(* IEC 61131-3 sources: OpenFactory/examples/openplc, 13 files *)

(* ---- batch-mix-heat.st ---- *)
(*
  OpenFactory example PLC program: batch-mix-heat (scenes/batch-mix-heat.yaml), the batch recipe
  of PLAN 3.3: fill two ingredients to a level each, heat to a temperature, hold.
  Target: OpenPLC v3 runtime (IEC 61131-3 Structured Text), talking to the OpenFactory simulator
  as a Modbus TCP Slave Device. Setup: docs/guides/openplc-quickstart.md, then
  docs/guides/batch-mix-heat.md for this scene.

  Training and demo use only. Not a safety-rated program and not a safety-rated simulation.

  Sequence of operations (one batch, then held); BATCH_STEP holds the active step
    0.  Idle: wait 1 s after power-up for the transmitters' first readings, then start a batch
        if the mixing tank is empty (level below 0.02 m).
    10. Fill water: open XV_01 until the level reaches 0.10 m.
    20. Fill syrup: open XV_02 until the level reaches 0.16 m (the recipe: 0.06 m of syrup on
        0.10 m of water, 37.5 % syrup by volume; each valve's 1 s close adds a little).
    30. Heat: the heater runs until the temperature reaches 50 C.
    40. Hold: the batch is ready (PL_READY_DO lit); the heater keeps it at 50 C, on below
        49.5 C and off at 50 C.
    Interlocks, in every step: the high level switch (LSH) closes both inlet valves, and the
    heater runs only while the level covers it (0.10 m and above).

  I/O map: Modbus addresses come from the scene's int16_scaled lockfile
  (scenes/batch-mix-heat.int16_scaled.modbus.yaml) and the exported I/O list CSV. OpenPLC places
  a Slave Device's points from address 100 onward, so a zero-based Modbus address N maps to
  %IX100.N, %QX100.N or %IW100+N.
*)
PROGRAM batch_mix_heat
  VAR
    (* Discrete inputs from the simulator (Modbus DI:0..3) *)
    TK_01_LSH_DI AT %IX100.0 : BOOL;    (* DI:0 Batch Mixing Tank - high level switch (LSH), 0.5 m *)
    XV_01_ZSC_DI AT %IX100.1 : BOOL;    (* DI:1 Mixing Tank Water Inlet Valve - closed limit (ZSC) *)
    XV_02_ZSC_DI AT %IX100.2 : BOOL;    (* DI:2 Mixing Tank Syrup Inlet Valve - closed limit (ZSC) *)
    SIM_HEARTBEAT_DI AT %IX100.3 : BOOL; (* DI:3 OpenFactory simulator heartbeat, 1 Hz; not used here, watch it for a sim-down watchdog *)
    (* Coils to the simulator (Modbus CO:0..3) *)
    HTR_01_ON_DO AT %QX100.0 : BOOL;    (* CO:0 Batch Mixing Tank Immersion Heater - on command *)
    PL_READY_DO AT %QX100.1 : BOOL;     (* CO:1 Batch Ready Pilot Light *)
    XV_01_OPEN_DO AT %QX100.2 : BOOL;   (* CO:2 Mixing Tank Water Inlet Valve - open command *)
    XV_02_OPEN_DO AT %QX100.3 : BOOL;   (* CO:3 Mixing Tank Syrup Inlet Valve - open command *)
    (* Input registers (Modbus IR:0..1) *)
    TK_01_LT_AI AT %IW100 : INT;        (* IR:0 Batch Mixing Tank Level Transmitter, 0 to 32767 = 0 to 0.6 m *)
    TK_01_TT_AI AT %IW101 : INT;        (* IR:1 Batch Mixing Tank Temperature Transmitter, 0 to 32767 = 0 to 100 C *)
  END_VAR
  VAR
    WATER_SP : REAL := 0.10;            (* level at which the water fill ends, m *)
    BATCH_SP : REAL := 0.16;            (* level at which the syrup fill ends, m *)
    EMPTY_LVL : REAL := 0.02;           (* below this the tank is empty and can start a batch, m *)
    TEMP_SP : REAL := 50.0;             (* batch temperature, C *)
    HOLD_DB : REAL := 0.5;              (* the heater restarts this far below TEMP_SP in the hold, C *)
    COVER_LVL : REAL := 0.10;           (* heater low-level permissive, m *)
    STARTUP_DELAY : TIME := T#1s;       (* until the transmitters' first readings *)
    STARTUP_TMR : TON;
    BATCH_STEP : INT := 0;              (* the active step: 0, 10, 20, 30, 40; not STEP, an IEC 61131-3 keyword *)
    HEAT : BOOL := FALSE;               (* heater demand before the permissive *)
    LEVEL_M : REAL;
    TEMP_C : REAL;
  END_VAR

  LEVEL_M := INT_TO_REAL(TK_01_LT_AI) * 0.6 / 32767.0;
  TEMP_C := INT_TO_REAL(TK_01_TT_AI) * 100.0 / 32767.0;
  STARTUP_TMR(IN := TRUE, PT := STARTUP_DELAY);

  (* Transitions, one per scan *)
  CASE BATCH_STEP OF
    0:  IF STARTUP_TMR.Q AND LEVEL_M < EMPTY_LVL THEN BATCH_STEP := 10; END_IF;
    10: IF LEVEL_M >= WATER_SP THEN BATCH_STEP := 20; END_IF;
    20: IF LEVEL_M >= BATCH_SP THEN BATCH_STEP := 30; END_IF;
    30: IF TEMP_C >= TEMP_SP THEN BATCH_STEP := 40; END_IF;
  END_CASE;

  (* Actions; the hold is a thermostat with a deadband *)
  IF BATCH_STEP = 30 THEN
    HEAT := TRUE;
  ELSIF BATCH_STEP = 40 THEN
    IF TEMP_C >= TEMP_SP THEN
      HEAT := FALSE;
    ELSIF TEMP_C < TEMP_SP - HOLD_DB THEN
      HEAT := TRUE;
    END_IF;
  ELSE
    HEAT := FALSE;
  END_IF;
  XV_01_OPEN_DO := (BATCH_STEP = 10) AND NOT TK_01_LSH_DI;
  XV_02_OPEN_DO := (BATCH_STEP = 20) AND NOT TK_01_LSH_DI;
  HTR_01_ON_DO := HEAT AND LEVEL_M >= COVER_LVL;
  PL_READY_DO := (BATCH_STEP = 40);
END_PROGRAM

CONFIGURATION Config0
  RESOURCE Res0 ON PLC
    TASK task0(INTERVAL := T#20ms, PRIORITY := 0);
    PROGRAM instance0 WITH task0 : batch_mix_heat;
  END_RESOURCE
END_CONFIGURATION

(* ---- buffer-and-release.st ---- *)
(*
  OpenFactory example PLC program: buffer-and-release (scenes/buffer-and-release.yaml), PLAN 2.7.
  Target: OpenPLC v3 runtime (IEC 61131-3 Structured Text), talking to the OpenFactory simulator
  as a Modbus TCP Slave Device. Setup: docs/guides/openplc-quickstart.md, then
  docs/guides/buffer-and-release.md for this scene.

  Training and demo use only. Not a safety-rated program and not a safety-rated simulation.

  Sequence of operations
    1. Run both belts. Hold STP_01 raised, so boxes queue nose to tail on the buffer belt.
    2. Enable the box emitter once both belts have reported running for 1 s.
    3. A batch is ready when PE_FULL (under the third queued box) has been blocked for 1.5 s, which
       a moving box (1 s in the beam at 0.3 m/s) cannot do, and the blade has been back up for at
       least 2 s since the last batch.
    4. Release: lower STP_01 and count PE_REL rising edges on the outfeed belt. The outfeed runs
       three times faster than the buffer, so each released box pulls a gap and the eye clears
       between boxes. At the third, raise the blade: the fourth box is still behind the blade line.

  Timing margin: when the third box of a batch reaches PE_REL, the fourth box's front is about
  0.10 m behind the blade line, 0.33 s at 0.3 m/s. OpenPLC sees the eye up to 100 ms late and
  writes the raise up to 100 ms later, which that margin covers. The blade holds parts from the
  moment it starts rising; a box already over the blade line passes.

  I/O map: Modbus addresses come from the scene's int16_scaled lockfile
  (scenes/buffer-and-release.int16_scaled.modbus.yaml) and the exported I/O list CSV. OpenPLC
  places a Slave Device's points from address 100 onward, so a zero-based Modbus address N maps
  to %IX100.N or %QX100.N. The scene has no analog tags, so both lockfiles give the same addresses.
*)
PROGRAM buffer_release
  VAR
    (* Discrete inputs from the simulator (Modbus DI:0..6) *)
    CONV_BUF_RUN_DI AT %IX100.0 : BOOL; (* DI:0 Buffer Belt Conveyor - running feedback *)
    CONV_OUT_RUN_DI AT %IX100.1 : BOOL; (* DI:1 Outfeed Belt Conveyor - running feedback *)
    PE_FULL_DI AT %IX100.2 : BOOL;      (* DI:2 Buffer Batch Ready Photo Eye - beam blocked *)
    PE_REL_DI AT %IX100.3 : BOOL;       (* DI:3 Outfeed Release Count Photo Eye - beam blocked *)
    STP_01_DN_DI AT %IX100.4 : BOOL;    (* DI:4 Buffer Release Stopper - lowered limit *)
    STP_01_UP_DI AT %IX100.5 : BOOL;    (* DI:5 Buffer Release Stopper - raised limit *)
    SIM_HEARTBEAT_DI AT %IX100.6 : BOOL; (* DI:6 OpenFactory simulator heartbeat, 1 Hz; not used here, watch it for a sim-down watchdog *)
    (* Coils to the simulator (Modbus CO:0..3) *)
    CONV_BUF_RUN_DO AT %QX100.0 : BOOL; (* CO:0 Buffer Belt Conveyor - run command *)
    CONV_OUT_RUN_DO AT %QX100.1 : BOOL; (* CO:1 Outfeed Belt Conveyor - run command *)
    EMT_01_EN_DO AT %QX100.2 : BOOL;    (* CO:2 Buffer Belt Box Source - enable *)
    STP_01_RAISE_DO AT %QX100.3 : BOOL; (* CO:3 Buffer Release Stopper - raise solenoid *)
  END_VAR
  VAR
    BATCH : INT := 3;                   (* boxes per release *)
    BELTS_OK_DELAY : TIME := T#1s;      (* run feedback must hold this long to feed boxes *)
    FULL_DELAY : TIME := T#1500ms;      (* a standing box, not a passing one, at PE_FULL *)
    PAUSE : TIME := T#2s;               (* blade up at least this long between batches *)
    BELTS_OK_TMR : TON;                 (* both belts running, debounced *)
    FULL_TMR : TON;                     (* a box stands under PE_FULL: three are queued *)
    PAUSE_TMR : TON;                    (* the blade has been back up PAUSE since the last batch *)
    PE_REL_RISE : R_TRIG;               (* a released box reaches PE_REL *)
    RELEASING : BOOL;                   (* a batch is on its way out *)
    RELEASED : INT;                     (* boxes counted out in this batch *)
  END_VAR

  (* 1. Belts run *)
  CONV_BUF_RUN_DO := TRUE;
  CONV_OUT_RUN_DO := TRUE;

  (* 2. Feed boxes only after both belts have reported running for BELTS_OK_DELAY *)
  BELTS_OK_TMR(IN := CONV_BUF_RUN_DI AND CONV_OUT_RUN_DI, PT := BELTS_OK_DELAY);
  EMT_01_EN_DO := BELTS_OK_TMR.Q;

  (* 3. A batch is ready: three queued, and the blade up long enough since the last batch *)
  FULL_TMR(IN := PE_FULL_DI, PT := FULL_DELAY);
  PAUSE_TMR(IN := STP_01_UP_DI AND NOT RELEASING, PT := PAUSE);
  IF FULL_TMR.Q AND PAUSE_TMR.Q AND NOT RELEASING THEN
    RELEASING := TRUE;
    RELEASED := 0;
  END_IF;

  (* 4. Count the batch out on the outfeed; raise the blade at the last one *)
  PE_REL_RISE(CLK := PE_REL_DI);
  IF PE_REL_RISE.Q AND RELEASING THEN
    RELEASED := RELEASED + 1;
    IF RELEASED >= BATCH THEN
      RELEASING := FALSE;
    END_IF;
  END_IF;
  STP_01_RAISE_DO := NOT RELEASING;
END_PROGRAM

CONFIGURATION Config0
  RESOURCE Res0 ON PLC
    TASK task0(INTERVAL := T#20ms, PRIORITY := 0);
    PROGRAM instance0 WITH task0 : buffer_release;
  END_RESOURCE
END_CONFIGURATION

(* ---- conveyor-start-stop.st ---- *)
(*
  OpenFactory example PLC program: conveyor-start-stop (scenes/conveyor-start-stop.yaml), the
  hello-world scene of PLAN 2.7.
  Target: OpenPLC v3 runtime (IEC 61131-3 Structured Text), talking to the OpenFactory simulator
  as a Modbus TCP Slave Device. Setup: docs/guides/openplc-quickstart.md, then
  docs/guides/conveyor-start-stop.md for this scene.

  Training and demo use only. Not a safety-rated program and not a safety-rated simulation.
  A real stop circuit is hard-wired; a PLC stop input like this one is an operator convenience.

  Sequence of operations
    1. Turning SS_01 to RUN starts the line: CONV_01 runs and stays running (seal-in) while SS_01
       stays in RUN and PB_STOP is not pressed. The scene starts with SS_01 in RUN, so the line
       starts on the first scan that sees it there.
    2. PB_STOP is wired normally closed (the scene binds it with invert: true): PB_STOP_DI is TRUE
       while the button is released, and a broken wire reads as a press, so it fails safe.
       Pressing it drops the seal-in. To restart, turn SS_01 to OFF and back to RUN.
    3. A selector reading OFF and RUN at once (a wiring fault) stops the line too.
    4. Once CONV_01 has reported running for 1 s, enable the box emitter EMT_01.
    5. PL_RUN shows the running feedback, not the command.
    Boxes ride the belt end to end and reach REM_01.

  I/O map: Modbus addresses come from the scene's int16_scaled lockfile
  (scenes/conveyor-start-stop.int16_scaled.modbus.yaml) and the exported I/O list CSV. OpenPLC
  places a Slave Device's points from address 100 onward, so a zero-based Modbus address N maps to
  %IX100.N or %QX100.N. This scene has no analog tags, so the float32 and int16_scaled lockfiles
  give the same addresses (ADR-0004 decision 8).

  Why the emitter waits 1 s: see examples/openplc/sorting-by-height.st. When OpenPLC (re)connects,
  its input image can hold old feedback for one poll, and an enable written straight from it can
  chatter and drop two boxes on top of each other.
*)
PROGRAM start_stop
  VAR
    (* Discrete inputs from the simulator (Modbus DI:0..4) *)
    CONV_01_RUN_DI AT %IX100.0 : BOOL;  (* DI:0 Transfer Belt Conveyor - running feedback *)
    PB_STOP_DI AT %IX100.1 : BOOL;      (* DI:1 Transfer Conveyor Stop Pushbutton - NC, TRUE = released *)
    SS_01_OFF_DI AT %IX100.2 : BOOL;    (* DI:2 Off/Run Selector Switch - in OFF *)
    SS_01_RUN_DI AT %IX100.3 : BOOL;    (* DI:3 Off/Run Selector Switch - in RUN *)
    SIM_HEARTBEAT_DI AT %IX100.4 : BOOL; (* DI:4 OpenFactory simulator heartbeat, 1 Hz; not used here, watch it for a sim-down watchdog *)
    (* Coils to the simulator (Modbus CO:0..2) *)
    CONV_01_RUN_DO AT %QX100.0 : BOOL;  (* CO:0 Transfer Belt Conveyor - run command *)
    EMT_01_EN_DO AT %QX100.1 : BOOL;    (* CO:1 Transfer Belt Box Source - enable *)
    PL_RUN_DO AT %QX100.2 : BOOL;       (* CO:2 Transfer Conveyor Running Pilot Light *)
  END_VAR
  VAR
    BELT_OK_DELAY : TIME := T#1s;       (* running feedback must hold this long to feed boxes *)
    BELT_OK_TMR : TON;                  (* belt running, debounced *)
    SS_RUN_RISE : R_TRIG;               (* selector turned to RUN (also the first scan in RUN) *)
    RUN_OK : BOOL;                      (* selector in RUN only, stop button released *)
    RUN_LATCH : BOOL;                   (* the line is started (seal-in) *)
  END_VAR

  (* 1-3. Start on a turn to RUN, seal in, drop on stop, OFF, or a selector wiring fault *)
  RUN_OK := SS_01_RUN_DI AND NOT SS_01_OFF_DI AND PB_STOP_DI;
  SS_RUN_RISE(CLK := SS_01_RUN_DI);
  RUN_LATCH := (SS_RUN_RISE.Q OR RUN_LATCH) AND RUN_OK;
  CONV_01_RUN_DO := RUN_LATCH;

  (* 4. Feed boxes only after the belt has reported running for BELT_OK_DELAY *)
  BELT_OK_TMR(IN := RUN_LATCH AND CONV_01_RUN_DI, PT := BELT_OK_DELAY);
  EMT_01_EN_DO := BELT_OK_TMR.Q;

  (* 5. Running light from feedback *)
  PL_RUN_DO := CONV_01_RUN_DI;
END_PROGRAM

CONFIGURATION Config0
  RESOURCE Res0 ON PLC
    TASK task0(INTERVAL := T#20ms, PRIORITY := 0);
    PROGRAM instance0 WITH task0 : start_stop;
  END_RESOURCE
END_CONFIGURATION

(* ---- inline-reject.st ---- *)
(*
  OpenFactory example PLC program: inline-reject (scenes/inline-reject.yaml).
  Target: OpenPLC v3 runtime (IEC 61131-3 Structured Text), talking to the OpenFactory simulator
  as a Modbus TCP Slave Device. Setup: docs/guides/openplc-quickstart.md.

  Training and demo use only. Not a safety-rated program and not a safety-rated simulation.

  The scene was built in the scene editor from `openfactory new`, without the file being opened
  (docs/guides/inline-reject.md). This program is a line-for-line port of the stand-in script,
  examples/pyplc/inline-reject.py.

  Sequence of operations
    1. Run both belt conveyors (CONV_01 feeds CONV_02 end to end).
    2. Enable the box emitter once both belts have reported running for 1 s without a break.
    3. PE_01 sits 0.3 m above CONV_02: oversize boxes (0.4 m) break the beam, good ones (0.2 m)
       pass under it. On each PE_01 rising edge, start that box's own REJECT_DELAY timer for its
       travel from the eye to the pusher plate, then extend CYL_01 when it expires; the plate
       pushes the box off the side of CONV_02 into the reject bin, REM_01. Each oversize box
       takes the next of four slots (a ring: REJECT_PEND_n and REJECT_TMR_n).
    4. Retract CYL_01 as soon as its extended limit (CYL_01_EXTENDED_DI) is made.
    Good boxes ride on to the end of CONV_02 and reach REM_02.

  I/O map: Modbus addresses come from the scene's lockfiles (scenes/inline-reject.*.modbus.yaml;
  this scene has no analog tags, so both give the same addresses). OpenPLC places a Slave
  Device's points from address 100 onward, so a zero-based Modbus address N maps to %IX100.N or
  %QX100.N.

  Timing: the eye and the plate are 1.0 m apart along CONV_02, as on sorting-by-height, so the
  box is due at the plate 2.08 s after it trips the eye at 0.5 m/s; REJECT_DELAY is 2.08 s minus
  OpenPLC's average 0.10 s polling latency, as the sorter's DIVERT_DELAY is.
*)
PROGRAM inline_reject
  VAR
    (* Discrete inputs from the simulator (Modbus DI:0..4) *)
    CONV_01_RUNNING_DI AT %IX100.0 : BOOL;  (* DI:0 Infeed Belt Conveyor - running feedback *)
    CONV_02_RUNNING_DI AT %IX100.1 : BOOL;  (* DI:1 Outfeed Belt Conveyor - running feedback *)
    CYL_01_EXTENDED_DI AT %IX100.2 : BOOL;  (* DI:2 Oversize Box Reject Pusher - extended limit *)
    PE_01_DI AT %IX100.3 : BOOL;            (* DI:3 Oversize Box Photo Eye - beam blocked *)
    SIM_HEARTBEAT_DI AT %IX100.4 : BOOL;    (* DI:4 OpenFactory simulator heartbeat, 1 Hz; not used here *)
    (* Coils to the simulator (Modbus CO:0..3) *)
    CONV_01_RUN_DO AT %QX100.0 : BOOL;      (* CO:0 Infeed Belt Conveyor - run command *)
    CONV_02_RUN_DO AT %QX100.1 : BOOL;      (* CO:1 Outfeed Belt Conveyor - run command *)
    CYL_01_EXTEND_DO AT %QX100.2 : BOOL;    (* CO:2 Oversize Box Reject Pusher - extend solenoid *)
    EMT_01_DO AT %QX100.3 : BOOL;           (* CO:3 Infeed Box Source - enable *)
  END_VAR
  VAR
    REJECT_DELAY : TIME := T#1980ms;    (* eye-to-plate travel, less average polling latency *)
    BELTS_OK_DELAY : TIME := T#1s;      (* run feedback must hold this long to feed boxes *)
    BELTS_OK_TMR : TON;                 (* both belts running, debounced *)
    PE_01_RISE : R_TRIG;                (* an oversize box arrives at PE_01 *)
    REJECT_TMR_0 : TON;                 (* eye-to-plate travel timer, slot 0 *)
    REJECT_TMR_1 : TON;                 (* eye-to-plate travel timer, slot 1 *)
    REJECT_TMR_2 : TON;                 (* eye-to-plate travel timer, slot 2 *)
    REJECT_TMR_3 : TON;                 (* eye-to-plate travel timer, slot 3 *)
    REJECT_PEND_0 : BOOL;               (* slot 0 holds an oversize box on its way to the pusher *)
    REJECT_PEND_1 : BOOL;               (* slot 1 holds an oversize box on its way to the pusher *)
    REJECT_PEND_2 : BOOL;               (* slot 2 holds an oversize box on its way to the pusher *)
    REJECT_PEND_3 : BOOL;               (* slot 3 holds an oversize box on its way to the pusher *)
    NEXT_SLOT : INT := 0;               (* ring index: the slot the next oversize box takes, 0..3 *)
    PUSH_CMD : BOOL;                    (* pusher extend request, held until the extended limit *)
  END_VAR

  (* 1. Belts run *)
  CONV_01_RUN_DO := TRUE;
  CONV_02_RUN_DO := TRUE;

  (* 2. Feed boxes only after both belts have reported running for BELTS_OK_DELAY *)
  BELTS_OK_TMR(IN := CONV_01_RUNNING_DI AND CONV_02_RUNNING_DI, PT := BELTS_OK_DELAY);
  EMT_01_DO := BELTS_OK_TMR.Q;

  (* 3. Oversize box at the eye: give it the next slot and its own travel timer *)
  PE_01_RISE(CLK := PE_01_DI);
  IF PE_01_RISE.Q THEN
    CASE NEXT_SLOT OF
      0: REJECT_PEND_0 := TRUE;
      1: REJECT_PEND_1 := TRUE;
      2: REJECT_PEND_2 := TRUE;
      3: REJECT_PEND_3 := TRUE;
    END_CASE;
    NEXT_SLOT := (NEXT_SLOT + 1) MOD 4;
  END_IF;

  (* 3a. Each slot's box is due at the plate: extend *)
  REJECT_TMR_0(IN := REJECT_PEND_0, PT := REJECT_DELAY);
  IF REJECT_TMR_0.Q THEN
    REJECT_PEND_0 := FALSE;
    PUSH_CMD := TRUE;
  END_IF;
  REJECT_TMR_1(IN := REJECT_PEND_1, PT := REJECT_DELAY);
  IF REJECT_TMR_1.Q THEN
    REJECT_PEND_1 := FALSE;
    PUSH_CMD := TRUE;
  END_IF;
  REJECT_TMR_2(IN := REJECT_PEND_2, PT := REJECT_DELAY);
  IF REJECT_TMR_2.Q THEN
    REJECT_PEND_2 := FALSE;
    PUSH_CMD := TRUE;
  END_IF;
  REJECT_TMR_3(IN := REJECT_PEND_3, PT := REJECT_DELAY);
  IF REJECT_TMR_3.Q THEN
    REJECT_PEND_3 := FALSE;
    PUSH_CMD := TRUE;
  END_IF;

  (* 4. Retract on the extended limit *)
  IF CYL_01_EXTENDED_DI THEN
    PUSH_CMD := FALSE;
  END_IF;
  CYL_01_EXTEND_DO := PUSH_CMD;
END_PROGRAM

CONFIGURATION Config0
  RESOURCE Res0 ON PLC
    TASK task0(INTERVAL := T#20ms, PRIORITY := 0);
    PROGRAM instance0 WITH task0 : inline_reject;
  END_RESOURCE
END_CONFIGURATION

(* ---- palletizer-lite.st ---- *)
(*
  OpenFactory example PLC program: palletizer-lite (scenes/palletizer-lite.yaml), PLAN 2.7.
  Target: OpenPLC v3 runtime (IEC 61131-3 Structured Text), talking to the OpenFactory simulator
  as a Modbus TCP Slave Device. Setup: docs/guides/openplc-quickstart.md, then
  docs/guides/palletizer-lite.md for this scene.

  Training and demo use only. Not a safety-rated program and not a safety-rated simulation.

  Sequence of operations
    1. Run both belts and hold both stoppers raised; enable the box source once both belts have
       reported running for 1 s. Boxes queue at STP_IN, the first one under the gantry.
    2. Pick and place, one box per cycle (the gantry has no raised switch, so each rise is timed):
       with a box at PE_PICK, the gantry at the pick side, fewer than LAYER_BOXES placed in this
       layer, and no layer leaving: PICK_STEP 1 lower, 2 grip, 3 rise, 4 traverse, 5 lower,
       6 release, 7 rise, 8 return, back to 0. (STEP is a reserved word in IEC 61131-3.) Count each box placed. The layer-forming belt carries it to
       the row queueing at STP_LYR.
    3. A layer is complete when LAYER_BOXES have been placed and PE_ROW (under the fourth queued
       box) has been blocked for 1 s, which a passing box (0.6 s in the beam) cannot do. Lower
       STP_LYR for LAYER_OUT to send the layer to the discharge, raise it, and start the count
       again. Counting placements, not just watching PE_ROW, keeps a fifth box from being set
       down while the row completes and riding out with the layer.

  I/O map: Modbus addresses come from the scene's int16_scaled lockfile
  (scenes/palletizer-lite.int16_scaled.modbus.yaml) and the exported I/O list CSV. OpenPLC places
  a Slave Device's points from address 100 onward, eight bits to a byte: zero-based Modbus address
  N maps to %IX(100 + N / 8).(N MOD 8), and likewise for %QX. The scene has no analog tags, so
  both lockfiles give the same addresses.
*)
PROGRAM palletizer
  VAR
    (* Discrete inputs from the simulator (Modbus DI:0..8) *)
    CONV_IN_RUN_DI AT %IX100.0 : BOOL;  (* DI:0 Palletizer Infeed Belt Conveyor - running *)
    CONV_LYR_RUN_DI AT %IX100.1 : BOOL; (* DI:1 Layer Forming Belt Conveyor - running *)
    PE_PICK_DI AT %IX100.2 : BOOL;      (* DI:2 Infeed Box At Pick Position Photo Eye *)
    PE_ROW_DI AT %IX100.3 : BOOL;       (* DI:3 Layer Row Complete Photo Eye *)
    PP_01_AT_PICK_DI AT %IX100.4 : BOOL;  (* DI:4 Transfer Gantry - at pick side *)
    PP_01_AT_PLACE_DI AT %IX100.5 : BOOL; (* DI:5 Transfer Gantry - at place side *)
    PP_01_DOWN_DI AT %IX100.6 : BOOL;   (* DI:6 Transfer Gantry - pad lowered *)
    PP_01_HOLD_DI AT %IX100.7 : BOOL;   (* DI:7 Transfer Gantry - holding a part *)
    SIM_HEARTBEAT_DI AT %IX100.8 : BOOL; (* DI:8 OpenFactory simulator heartbeat, 1 Hz; not used here, watch it for a sim-down watchdog *)
    (* Coils to the simulator (Modbus CO:0..7) *)
    CONV_IN_RUN_DO AT %QX100.0 : BOOL;  (* CO:0 Palletizer Infeed Belt Conveyor - run *)
    CONV_LYR_RUN_DO AT %QX100.1 : BOOL; (* CO:1 Layer Forming Belt Conveyor - run *)
    EMT_01_EN_DO AT %QX100.2 : BOOL;    (* CO:2 Palletizer Infeed Box Source - enable *)
    PP_01_GRIP_DO AT %QX100.3 : BOOL;   (* CO:3 Transfer Gantry - grip *)
    PP_01_LOWER_DO AT %QX100.4 : BOOL;  (* CO:4 Transfer Gantry - lower pad *)
    PP_01_TRAV_DO AT %QX100.5 : BOOL;   (* CO:5 Transfer Gantry - traverse to place side *)
    STP_IN_RAISE_DO AT %QX100.6 : BOOL; (* CO:6 Infeed Pick Position Stopper - raise *)
    STP_LYR_RAISE_DO AT %QX100.7 : BOOL; (* CO:7 Layer Forming Stopper - raise *)
  END_VAR
  VAR
    LAYER_BOXES : INT := 4;             (* boxes per layer *)
    BELTS_OK_DELAY : TIME := T#1s;      (* run feedback must hold this long to feed boxes *)
    RISE : TIME := T#400ms;             (* pad rise, lower_time_s 0.3 plus margin *)
    SETTLE : TIME := T#200ms;           (* the released box drops onto the belt *)
    ROW_DELAY : TIME := T#1s;           (* a standing box, not a passing one, at PE_ROW *)
    LAYER_OUT : TIME := T#3s;           (* four boxes (1.2 m) clear the blade at 0.5 m/s *)
    BELTS_OK_TMR : TON;                 (* both belts running, debounced *)
    RISE_TMR : TON;                     (* the pad has had time to rise *)
    SETTLE_TMR : TON;                   (* the released box has settled on the belt *)
    ROW_TMR : TON;                      (* a box stands under PE_ROW *)
    LAYER_TMR : TON;                    (* the layer has had time to leave *)
    PICK_STEP : INT := 0;               (* pick-and-place step, 0 = waiting at the pick side *)
    LAYER_OUT_ON : BOOL;                (* a layer is leaving *)
    PLACED : INT := 0;                  (* boxes placed in the layer being formed *)
  END_VAR

  (* 1. Belts run; stoppers hold; feed boxes once both belts report running for 1 s *)
  CONV_IN_RUN_DO := TRUE;
  CONV_LYR_RUN_DO := TRUE;
  STP_IN_RAISE_DO := TRUE;
  BELTS_OK_TMR(IN := CONV_IN_RUN_DI AND CONV_LYR_RUN_DI, PT := BELTS_OK_DELAY);
  EMT_01_EN_DO := BELTS_OK_TMR.Q;

  (* 2. Pick and place, one box per cycle; the timers run only in the steps that use them *)
  RISE_TMR(IN := PICK_STEP = 3 OR PICK_STEP = 7, PT := RISE);
  SETTLE_TMR(IN := PICK_STEP = 6 AND NOT PP_01_HOLD_DI, PT := SETTLE);
  CASE PICK_STEP OF
    0: IF PE_PICK_DI AND PP_01_AT_PICK_DI AND PLACED < LAYER_BOXES AND NOT LAYER_OUT_ON THEN
         PICK_STEP := 1;
       END_IF;
    1: IF PP_01_DOWN_DI THEN PICK_STEP := 2; END_IF;
    2: IF PP_01_HOLD_DI THEN PICK_STEP := 3; END_IF;
    3: IF RISE_TMR.Q THEN PICK_STEP := 4; END_IF;
    4: IF PP_01_AT_PLACE_DI THEN PICK_STEP := 5; END_IF;
    5: IF PP_01_DOWN_DI THEN PICK_STEP := 6; END_IF;
    6: IF SETTLE_TMR.Q THEN
         PICK_STEP := 7;
         PLACED := PLACED + 1;
       END_IF;
    7: IF RISE_TMR.Q THEN PICK_STEP := 8; END_IF;
    8: IF PP_01_AT_PICK_DI THEN PICK_STEP := 0; END_IF;
  END_CASE;
  PP_01_LOWER_DO := PICK_STEP = 1 OR PICK_STEP = 2 OR PICK_STEP = 5 OR PICK_STEP = 6;
  PP_01_GRIP_DO := PICK_STEP = 2 OR PICK_STEP = 3 OR PICK_STEP = 4 OR PICK_STEP = 5;
  PP_01_TRAV_DO := PICK_STEP = 4 OR PICK_STEP = 5 OR PICK_STEP = 6 OR PICK_STEP = 7;

  (* 3. A complete row leaves as one layer *)
  ROW_TMR(IN := PE_ROW_DI, PT := ROW_DELAY);
  IF ROW_TMR.Q AND PLACED >= LAYER_BOXES AND NOT LAYER_OUT_ON THEN
    LAYER_OUT_ON := TRUE;
  END_IF;
  LAYER_TMR(IN := LAYER_OUT_ON, PT := LAYER_OUT);
  IF LAYER_TMR.Q THEN
    LAYER_OUT_ON := FALSE;
    PLACED := 0;
  END_IF;
  STP_LYR_RAISE_DO := NOT LAYER_OUT_ON;
END_PROGRAM

CONFIGURATION Config0
  RESOURCE Res0 ON PLC
    TASK task0(INTERVAL := T#20ms, PRIORITY := 0);
    PROGRAM instance0 WITH task0 : palletizer;
  END_RESOURCE
END_CONFIGURATION

(* ---- plantpax-tank-level.st ---- *)
(*
  OpenFactory example PLC program: plantpax-tank-level (scenes/plantpax-tank-level.yaml), the
  PlantPAx demo plant of PLAN 3.4 controlled without PlantPAx: tank-level-pid's level loop closed
  with OpenPLC's PID function block, plus the transfer pump. The PlantPAx version of the same
  control is the L5X from `openfactory export ... --format plantpax` (docs/plantpax.md).
  Target: OpenPLC v3 runtime (IEC 61131-3 Structured Text), talking to the OpenFactory simulator
  as a Modbus TCP Slave Device. Setup: docs/guides/openplc-quickstart.md, then
  docs/guides/plantpax-tank-level.md for this scene.

  Training and demo use only. Not a safety-rated program and not a safety-rated simulation.

  The PID block is the one in OpenPLC's compiler library (matiec lib/pid_st.txt, from the IEC
  61131-3 2nd edition draft): XOUT := KP * (ERROR + ITERM.XOUT / TR + DTERM.XOUT * TD) with
  ERROR := PV - SP. The error is PV minus SP, so a loop that opens the inlet valve on a low level
  needs a negative KP. Its integral (lib/integral_st.txt) is a rectangular sum of ERROR times
  TIME_TO_REAL(CYCLE). It has no output limit and no anti-windup: LIMIT clamps the output here,
  and the interlock holds the block in manual so it cannot wind up while overridden.
  [TBD: verify on the first OpenPLC run] that TIME_TO_REAL(T#20ms) is 0.02 (seconds) in the
  runtime; the gains below assume seconds, as the stand-in script does.

  Sequence of operations
    1. Read the level from the transmitter, raw 0 to 32767 for 0 to 2 m.
    2. PI control: the valve position is KP * (e + sum(e * 0.02 s) / TR) with e = level - 1.0 m.
    3. The output is limited to 0 to 100 % and written to the valve, raw 0 to 32767.
    4. Interlock: while the high level switch (LSH) is on, the valve is closed and the PID is
       held in manual at 0 % (no windup while it is overridden).
    5. For the first second the PID runs in manual at the valve's starting position (66 %),
       tracking the level, then switches to automatic bumplessly: the level input reads 0 until
       its first poll, and starting in automatic on that would slam the valve shut.
    6. The transfer pump P_01 starts 20 s after power-up (the demo's load step) and runs while
       the low level switch (LSL) is off: LSL is its interlock against running the tank dry.

  I/O map: Modbus addresses come from the scene's int16_scaled lockfile
  (scenes/plantpax-tank-level.int16_scaled.modbus.yaml) and the exported I/O list CSV. OpenPLC places
  a Slave Device's points from address 100 onward, so a zero-based Modbus address N maps to
  %IX100.N, %IW100+N, or %QW100+N.
*)
PROGRAM plantpax_tank
  VAR
    (* Discrete inputs from the simulator (Modbus DI:0..3) *)
    P_01_RUN_DI AT %IX100.0 : BOOL;     (* DI:0 Level Control Tank Transfer Pump - running feedback *)
    TK_01_LSH_DI AT %IX100.1 : BOOL;    (* DI:1 Level Control Tank - high level switch (LSH), 1.8 m *)
    TK_01_LSL_DI AT %IX100.2 : BOOL;    (* DI:2 Level Control Tank - low level switch (LSL), 0.3 m *)
    SIM_HEARTBEAT_DI AT %IX100.3 : BOOL; (* DI:3 OpenFactory simulator heartbeat, 1 Hz; not used here, watch it for a sim-down watchdog *)
    (* Coils to the simulator (Modbus CO:0) *)
    P_01_RUN_DO AT %QX100.0 : BOOL;     (* CO:0 Level Control Tank Transfer Pump - run command *)
    (* Input registers (Modbus IR:0..1) *)
    FV_01_ZT_AI AT %IW100 : INT;        (* IR:0 Tank Inlet Level Control Valve - position feedback, 0 to 32767 = 0 to 100 % *)
    TK_01_LT_AI AT %IW101 : INT;        (* IR:1 Level Control Tank Level Transmitter, 0 to 32767 = 0 to 2 m *)
    (* Holding registers to the simulator (Modbus HR:0) *)
    FV_01_POS_AO AT %QW100 : INT;       (* HR:0 Tank Inlet Level Control Valve - position command, 0 to 32767 = 0 to 100 % *)
  END_VAR
  VAR
    SP : REAL := 1.0;                   (* level setpoint, m *)
    KP : REAL := -400.0;                (* % per m; negative: the PID's error is PV - SP *)
    TR : REAL := 6.0;                   (* reset time, s *)
    START_PCT : REAL := 66.0;           (* valve position at start, % *)
    STARTUP_DELAY : TIME := T#1s;       (* manual until the level reading is live *)
    STARTUP_TMR : TON;
    LOAD_DELAY : TIME := T#20s;         (* the transfer pump starts: the demo's load step *)
    LOAD_TMR : TON;
    LIC : PID;                          (* the level controller *)
    LEVEL_M : REAL;
    MANUAL_X0 : REAL;
    OUT_PCT : REAL;
  END_VAR

  (* 1. Level in metres *)
  LEVEL_M := INT_TO_REAL(TK_01_LT_AI) * 2.0 / 32767.0;

  (* 5. Manual at the starting position until the startup delay is done *)
  STARTUP_TMR(IN := TRUE, PT := STARTUP_DELAY);
  IF STARTUP_TMR.Q THEN
    MANUAL_X0 := 0.0;
  ELSE
    MANUAL_X0 := START_PCT / KP;         (* in manual the block outputs KP * X0 *)
  END_IF;

  (* 2. PI on the level; 4. held in manual at 0 % while the high switch overrides it *)
  LIC(AUTO := STARTUP_TMR.Q AND NOT TK_01_LSH_DI, PV := LEVEL_M, SP := SP, X0 := MANUAL_X0,
      KP := KP, TR := TR, TD := 0.0, CYCLE := T#20ms);

  (* 3. Limit to the valve's range; 4. the interlock closes it *)
  IF TK_01_LSH_DI THEN
    OUT_PCT := 0.0;
  ELSE
    OUT_PCT := LIMIT(0.0, LIC.XOUT, 100.0);
  END_IF;
  FV_01_POS_AO := REAL_TO_INT(OUT_PCT * 32767.0 / 100.0);

  (* 6. The transfer pump: started 20 s after power-up, interlocked off by the low level switch *)
  LOAD_TMR(IN := TRUE, PT := LOAD_DELAY);
  P_01_RUN_DO := LOAD_TMR.Q AND NOT TK_01_LSL_DI;
END_PROGRAM

CONFIGURATION Config0
  RESOURCE Res0 ON PLC
    TASK task0(INTERVAL := T#20ms, PRIORITY := 0);
    PROGRAM instance0 WITH task0 : plantpax_tank;
  END_RESOURCE
END_CONFIGURATION

(* ---- silo-batch-weigh.st ---- *)
(*
  OpenFactory example PLC program: silo-batch-weigh (scenes/silo-batch-weigh.yaml), the bulk
  solids scene of PLAN 5.7a: an airlock and a screw fill a weigh hopper to a batch weight, then a
  gate empties it into a mixer; the silo refills itself through its roof gate.
  Target: OpenPLC v3 runtime (IEC 61131-3 Structured Text), talking to the OpenFactory simulator
  as a Modbus TCP Slave Device. Setup: docs/guides/openplc-quickstart.md, then
  docs/guides/silo-batch-weigh.md for this scene. A port of examples/pyplc/silo-batch-weigh.py:
  same sequence, same tag names.

  Training and demo use only. Not a safety-rated program and not a safety-rated simulation.

  Sequence of operations; BATCH_STEP holds the active step
    Silo refill, on its own: SG_01 opens when the silo's net weight falls below REFILL_ON_KG and
    closes above REFILL_OFF_KG.
    1. FAST (10): the screw runs and the airlock turns at 100 % until the hopper's net weight
       reaches TARGET_KG - FAST_PREACT_KG (the screw runs full: 50 kg is still on it).
    2. SLOW (20): the airlock turns at SLOW_PCT until the net weight reaches
       TARGET_KG - SLOW_PREACT_KG (what the screw carries at that rate in its travel time).
    3. EMPTYING (30): the airlock stops; the screw runs on for SCREW_RUN_ON, then stops.
    4. DISCHARGE (40): the hopper's gate SG_02 opens until the hopper is empty.
    5. CLOSING (50): when the gate's closed limit switch is made, the next batch starts.
    The airlock runs only while the screw runs and is not plugged.

  I/O map: Modbus addresses come from the scene's int16_scaled lockfile
  (scenes/silo-batch-weigh.int16_scaled.modbus.yaml) and the exported I/O list CSV. OpenPLC
  places a Slave Device's points from address 100 onward, eight bits a byte: a zero-based
  discrete address N maps to %IX(100 + N / 8).(N mod 8), a register N to %IW100+N.
*)
PROGRAM silo_batch_weigh
  VAR
    (* Discrete inputs from the simulator (Modbus DI:0..12) *)
    RV_01_PLUG_DI AT %IX100.0 : BOOL;   (* DI:0 Silo Discharge Rotary Airlock - plug switch *)
    RV_01_RUN_DI AT %IX100.1 : BOOL;    (* DI:1 Silo Discharge Rotary Airlock - running *)
    SC_01_PLUG_DI AT %IX100.2 : BOOL;   (* DI:2 Weigh Hopper Feed Screw Conveyor - plug switch *)
    SC_01_RUN_DI AT %IX100.3 : BOOL;    (* DI:3 Weigh Hopper Feed Screw Conveyor - running *)
    SC_01_ZSS_DI AT %IX100.4 : BOOL;    (* DI:4 Weigh Hopper Feed Screw Conveyor - zero-speed switch *)
    SG_01_ZSC_DI AT %IX100.5 : BOOL;    (* DI:5 Silo Fill Gate - closed limit (ZSC) *)
    SG_01_ZSO_DI AT %IX100.6 : BOOL;    (* DI:6 Silo Fill Gate - open limit (ZSO) *)
    SG_02_ZSC_DI AT %IX100.7 : BOOL;    (* DI:7 Weigh Hopper Discharge Gate - closed limit (ZSC) *)
    SG_02_ZSO_DI AT %IX101.0 : BOOL;    (* DI:8 Weigh Hopper Discharge Gate - open limit (ZSO) *)
    SILO_01_LSH_DI AT %IX101.1 : BOOL;  (* DI:9 Flour Storage Silo - high level switch (LSH) *)
    SILO_01_LSL_DI AT %IX101.2 : BOOL;  (* DI:10 Flour Storage Silo - low level switch (LSL) *)
    WH_01_LSH_DI AT %IX101.3 : BOOL;    (* DI:11 Batch Weigh Hopper - high level switch (LSH) *)
    SIM_HEARTBEAT_DI AT %IX101.4 : BOOL; (* DI:12 OpenFactory simulator heartbeat, 1 Hz; not used here, watch it for a sim-down watchdog *)
    (* Coils to the simulator (Modbus CO:0..3) *)
    RV_01_RUN_DO AT %QX100.0 : BOOL;    (* CO:0 Silo Discharge Rotary Airlock - run *)
    SC_01_RUN_DO AT %QX100.1 : BOOL;    (* CO:1 Weigh Hopper Feed Screw Conveyor - run *)
    SG_01_OPEN_DO AT %QX100.2 : BOOL;   (* CO:2 Silo Fill Gate - open (held) *)
    SG_02_OPEN_DO AT %QX100.3 : BOOL;   (* CO:3 Weigh Hopper Discharge Gate - open (held) *)
    (* Input registers (Modbus IR:0..2) *)
    SILO_01_LT_AI AT %IW100 : INT;      (* IR:0 Flour Storage Silo level, 0 to 32767 = 0 to 4.5 m *)
    SILO_01_WT_AI AT %IW101 : INT;      (* IR:1 Flour Storage Silo weight, 0 to 32767 = 0 to 10000 kg *)
    WH_01_WT_AI AT %IW102 : INT;        (* IR:2 Batch Weigh Hopper weight, 0 to 32767 = 0 to 750 kg *)
    (* Holding registers (Modbus HR:0) *)
    RV_01_SPD_AO AT %QW100 : INT;       (* HR:0 Silo Discharge Rotary Airlock speed, 0 to 32767 = 0 to 100 % *)
  END_VAR
  VAR
    SILO_TARE_KG : REAL := 1800.0;
    HOPPER_TARE_KG : REAL := 180.0;
    REFILL_ON_KG : REAL := 3500.0;
    REFILL_OFF_KG : REAL := 4500.0;
    TARGET_KG : REAL := 250.0;
    FAST_PREACT_KG : REAL := 65.0;      (* the screw's load running full (10 kg/s x 5 s) and a margin *)
    SLOW_PCT : REAL := 20.0;            (* 12 kg/s x 20 % = 2.4 kg/s *)
    SLOW_PREACT_KG : REAL := 12.0;      (* 2.4 kg/s x 5 s on the screw *)
    SCREW_RUN_ON : TIME := T#6s;        (* its travel time, 5 s, and a margin *)
    EMPTY_KG : REAL := 0.5;
    RUN_ON_TMR : TON;
    BATCH_STEP : INT := 10;             (* 10 FAST, 20 SLOW, 30 EMPTYING, 40 DISCHARGE, 50 CLOSING *)
    REFILL : BOOL := FALSE;
    SCREW_OK : BOOL;
    SILO_KG : REAL;
    NET_KG : REAL;
    SPEED_PCT : REAL;
  END_VAR

  SILO_KG := INT_TO_REAL(SILO_01_WT_AI) * 10000.0 / 32767.0 - SILO_TARE_KG;
  REFILL := (SILO_KG < REFILL_ON_KG OR REFILL) AND SILO_KG < REFILL_OFF_KG;
  SG_01_OPEN_DO := REFILL;

  NET_KG := INT_TO_REAL(WH_01_WT_AI) * 750.0 / 32767.0 - HOPPER_TARE_KG;
  SCREW_OK := SC_01_RUN_DI AND NOT SC_01_PLUG_DI;
  RUN_ON_TMR(IN := (BATCH_STEP = 30), PT := SCREW_RUN_ON);

  (* Transitions, one per scan *)
  CASE BATCH_STEP OF
    10: IF NET_KG >= TARGET_KG - FAST_PREACT_KG THEN BATCH_STEP := 20; END_IF;
    20: IF NET_KG >= TARGET_KG - SLOW_PREACT_KG THEN BATCH_STEP := 30; END_IF;
    30: IF RUN_ON_TMR.Q THEN BATCH_STEP := 40; END_IF;
    40: IF NET_KG <= EMPTY_KG THEN BATCH_STEP := 50; END_IF;
    50: IF SG_02_ZSC_DI THEN BATCH_STEP := 10; END_IF;
  END_CASE;

  (* Actions *)
  SC_01_RUN_DO := (BATCH_STEP = 10) OR (BATCH_STEP = 20) OR (BATCH_STEP = 30);
  RV_01_RUN_DO := ((BATCH_STEP = 10) OR (BATCH_STEP = 20)) AND SCREW_OK;
  IF BATCH_STEP = 10 THEN
    SPEED_PCT := 100.0;
  ELSE
    SPEED_PCT := SLOW_PCT;
  END_IF;
  RV_01_SPD_AO := REAL_TO_INT(SPEED_PCT * 32767.0 / 100.0);
  SG_02_OPEN_DO := (BATCH_STEP = 40);
END_PROGRAM

CONFIGURATION Config0
  RESOURCE Res0 ON PLC
    TASK task0(INTERVAL := T#20ms, PRIORITY := 0);
    PROGRAM instance0 WITH task0 : silo_batch_weigh;
  END_RESOURCE
END_CONFIGURATION

(* ---- sorting-by-color.st ---- *)
(*
  OpenFactory example PLC program: sorting-by-color (scenes/sorting-by-color.yaml), PLAN 2.7.
  Target: OpenPLC v3 runtime (IEC 61131-3 Structured Text), talking to the OpenFactory simulator
  as a Modbus TCP Slave Device. Setup: docs/guides/openplc-quickstart.md, then
  docs/guides/sorting-by-color.md for this scene.

  Training and demo use only. Not a safety-rated program and not a safety-rated simulation.

  Sequence of operations
    1. Run both belts; enable the box source once both have reported running for 1 s.
    2. On each CS_01_RED_DI rising edge (a red box under the color sensor), start that box's
       EXTEND_DELAY timer. When it expires, count the box as on its way to the arm: the arm
       extends while any red box is on its way. The delay lets a blue box already past the
       sensor clear the arm before it swings out (a swinging arm sweeps whatever it reaches).
    3. Each PE_RED rising edge (a red box arriving on the side lane) counts one red box off; the
       arm retracts when none is left on its way.
    Boxes are at least 4 s (2 m) apart, so one pending timer is enough; closer boxes would need a
    ring of timers as in examples/openplc/sorting-by-height.st.

  Timing: a red box is under the sensor for 0.6 s (0.3 m at 0.5 m/s), three OpenPLC polls. After
  EXTEND_DELAY (1.5 s) it is 0.75 m past the sensor and 0.85 m from the arm, which needs 0.5 s
  to swing out; the box ahead of it, at least 2 m ahead, is already past the arm's tip.

  I/O map: Modbus addresses come from the scene's int16_scaled lockfile
  (scenes/sorting-by-color.int16_scaled.modbus.yaml) and the exported I/O list CSV. OpenPLC places
  a Slave Device's points from address 100 onward, so a zero-based Modbus address N maps to
  %IX100.N or %QX100.N. The scene has no analog tags, so both lockfiles give the same addresses.
*)
PROGRAM color_sort
  VAR
    (* Discrete inputs from the simulator (Modbus DI:0..7) *)
    CONV_01_RUN_DI AT %IX100.0 : BOOL;  (* DI:0 Sorting Line Belt Conveyor - running *)
    CONV_RED_RUN_DI AT %IX100.1 : BOOL; (* DI:1 Red Box Lane Belt Conveyor - running *)
    CS_01_PART_DI AT %IX100.2 : BOOL;   (* DI:2 Red Box Color Sensor - part in range *)
    CS_01_RED_DI AT %IX100.3 : BOOL;    (* DI:3 Red Box Color Sensor - red seen *)
    DIV_01_EXT_DI AT %IX100.4 : BOOL;   (* DI:4 Red Box Divert Arm - extended limit *)
    DIV_01_RET_DI AT %IX100.5 : BOOL;   (* DI:5 Red Box Divert Arm - retracted limit *)
    PE_RED_DI AT %IX100.6 : BOOL;       (* DI:6 Red Box Lane Arrival Photo Eye *)
    SIM_HEARTBEAT_DI AT %IX100.7 : BOOL; (* DI:7 OpenFactory simulator heartbeat, 1 Hz; not used here, watch it for a sim-down watchdog *)
    (* Coils to the simulator (Modbus CO:0..3) *)
    CONV_01_RUN_DO AT %QX100.0 : BOOL;  (* CO:0 Sorting Line Belt Conveyor - run *)
    CONV_RED_RUN_DO AT %QX100.1 : BOOL; (* CO:1 Red Box Lane Belt Conveyor - run *)
    DIV_01_EXT_DO AT %QX100.2 : BOOL;   (* CO:2 Red Box Divert Arm - extend solenoid *)
    EMT_01_EN_DO AT %QX100.3 : BOOL;    (* CO:3 Sorting Line Box Source - enable *)
  END_VAR
  VAR
    BELTS_OK_DELAY : TIME := T#1s;      (* run feedback must hold this long to feed boxes *)
    EXTEND_DELAY : TIME := T#1500ms;    (* the red box is then 0.75 m past the sensor *)
    BELTS_OK_TMR : TON;                 (* both belts running, debounced *)
    EXTEND_TMR : TON;                   (* a red box's travel from the sensor toward the arm *)
    RED_RISE : R_TRIG;                  (* a red box arrives under the color sensor *)
    LANE_RISE : R_TRIG;                 (* a red box arrives on the side lane *)
    PENDING : BOOL;                     (* a red box is between the sensor and the extend point *)
    RED_OUT : INT := 0;                 (* red boxes between the extend point and the side lane *)
  END_VAR

  (* 1. Belts run; feed boxes once both report running for 1 s *)
  CONV_01_RUN_DO := TRUE;
  CONV_RED_RUN_DO := TRUE;
  BELTS_OK_TMR(IN := CONV_01_RUN_DI AND CONV_RED_RUN_DI, PT := BELTS_OK_DELAY);
  EMT_01_EN_DO := BELTS_OK_TMR.Q;

  (* 2. A red box at the sensor: after EXTEND_DELAY it is on its way to the arm *)
  RED_RISE(CLK := CS_01_RED_DI);
  IF RED_RISE.Q THEN
    PENDING := TRUE;
  END_IF;
  EXTEND_TMR(IN := PENDING, PT := EXTEND_DELAY);
  IF EXTEND_TMR.Q THEN
    PENDING := FALSE;
    RED_OUT := RED_OUT + 1;
  END_IF;

  (* 3. A red box on the side lane is done *)
  LANE_RISE(CLK := PE_RED_DI);
  IF LANE_RISE.Q AND RED_OUT > 0 THEN
    RED_OUT := RED_OUT - 1;
  END_IF;
  DIV_01_EXT_DO := RED_OUT > 0;
END_PROGRAM

CONFIGURATION Config0
  RESOURCE Res0 ON PLC
    TASK task0(INTERVAL := T#20ms, PRIORITY := 0);
    PROGRAM instance0 WITH task0 : color_sort;
  END_RESOURCE
END_CONFIGURATION

(* ---- sorting-by-height.st ---- *)
(*
  OpenFactory example PLC program: sorting-by-height (scenes/sorting-by-height.yaml).
  Target: OpenPLC v3 runtime (IEC 61131-3 Structured Text), talking to the OpenFactory simulator
  as a Modbus TCP Slave Device. Setup: docs/guides/openplc-quickstart.md.

  Training and demo use only. Not a safety-rated program and not a safety-rated simulation.

  Sequence of operations
    1. Run both belt conveyors (CONV_01 infeed, CONV_02 divert lane) and write both speed
       references, 100 % each.
    2. Enable the box emitter once both belts have reported running for 1 s without a break.
    3. PE_01 sits 0.3 m above the belt: tall boxes (0.4 m) break the beam, short ones (0.2 m) pass
       under it. On each PE_01 rising edge, start that box's own DIVERT_DELAY timer for its travel
       from the eye to the pusher plate, then extend CYL_01 when it expires. Each tall box takes
       the next of four divert slots (a ring: DIVERT_PEND_n and DIVERT_TMR_n), so a second tall
       box tripping the eye before the first is pushed keeps its own divert.
    4. Retract CYL_01 as soon as its extended limit (CYL_01_EXT_DI) is made.
    Tall boxes end up on CONV_02 and reach REM_02; short boxes stay on CONV_01 and reach REM_01.

  I/O map: Modbus addresses come from the scene's int16_scaled lockfile
  (scenes/sorting-by-height.int16_scaled.modbus.yaml) and the exported I/O list CSV
  (openfactory export ... --analog-encoding int16_scaled). OpenPLC places a Slave Device's points
  from address 100 onward, so a zero-based Modbus address N maps to %IX100.N, %QX100.N, or %QW100+N.
  Digital addresses (DI, CO) are identical in the float32 and int16_scaled lockfiles (ADR-0004
  decision 8); only the holding registers differ (float32 uses two per tag).

  Timing: PE_01 trips when a tall box's leading edge reaches x = 1.5 m; the plate starts pushing
  best when the box center is near x = 2.39 m, 2.08 s later at 0.5 m/s (the headless sorter test,
  tests/unit/test_sorter_headless.py). OpenPLC polls the simulator every 100 ms (Settings, Slave
  polling period), so the eye is seen up to 100 ms late and the extend coil written up to 100 ms
  late, about 100 ms on average; DIVERT_DELAY is 2.08 s minus that 0.10 s. A tall box blocks the
  beam for 0.6 s, well above the ~200 ms minimum pulse that 100 ms polling can catch.

  Divert queue: boxes are 0.3 m long at 0.5 m/s, so tall boxes can trip the eye about 0.8 s apart
  at the closest (box plus a gap that clears the beam), and up to three can be between the eye and
  the plate at once. Four slots cover that. A fifth box in transit would find its slot still busy:
  DIVERT_OVERRUN latches TRUE (watch it in the OpenPLC monitor) and that box is not diverted. The
  pusher needs 0.8 s to extend and retract, so tall boxes closer than that cannot all be pushed
  whatever the program does. tests/scenes/sorter-tall-pairs.yaml (every box tall, 1.5 s apart)
  exercises two pending diverts at once.

  Why the emitter waits 1 s: the emitter spawns a box the moment it is enabled. When OpenPLC
  (re)connects, its input image can still hold old feedback for one poll, so an enable written
  straight from the run feedback chatters on, off, on within ~0.3 s and drops two boxes on top of
  each other; the pusher then diverts both, short box included (seen in the first 1.14 run). The
  BELTS_OK_TMR permissive delay filters that out.
*)
PROGRAM sorter
  VAR
    (* Discrete inputs from the simulator (Modbus DI:0..5, same in every encoding) *)
    CONV_01_RUN_DI AT %IX100.0 : BOOL;  (* DI:0 Infeed Belt Conveyor - running feedback *)
    CYL_01_EXT_DI AT %IX100.1 : BOOL;   (* DI:1 Tall Box Divert Pusher - extended limit *)
    CYL_01_RET_DI AT %IX100.2 : BOOL;   (* DI:2 Tall Box Divert Pusher - retracted limit *)
    PE_01_DI AT %IX100.3 : BOOL;        (* DI:3 Infeed Tall Box Photo Eye - beam blocked *)
    CONV_02_RUN_DI AT %IX100.4 : BOOL;  (* DI:4 Divert Lane Belt Conveyor - running feedback *)
    SIM_HEARTBEAT_DI AT %IX100.5 : BOOL; (* DI:5 OpenFactory simulator heartbeat, 1 Hz; not used here, watch it for a sim-down watchdog *)
    (* Coils to the simulator (Modbus CO:0..3, same in every encoding) *)
    CONV_01_RUN_DO AT %QX100.0 : BOOL;  (* CO:0 Infeed Belt Conveyor - run command *)
    CYL_01_EXT_DO AT %QX100.1 : BOOL;   (* CO:1 Tall Box Divert Pusher - extend solenoid *)
    EMT_01_EN_DO AT %QX100.2 : BOOL;    (* CO:2 Infeed Box Source - enable *)
    CONV_02_RUN_DO AT %QX100.3 : BOOL;  (* CO:3 Divert Lane Belt Conveyor - run command *)
    (* Holding registers to the simulator (Modbus HR:0..1), int16_scaled: 0..32767 = 0..100 % *)
    CONV_01_SPD_AO AT %QW100 : INT;     (* HR:0 Infeed Belt Conveyor - speed command *)
    CONV_02_SPD_AO AT %QW101 : INT;     (* HR:1 Divert Lane Belt Conveyor - speed command *)
  END_VAR
  VAR
    SPEED_RAW : INT := 32767;           (* 100 % speed reference, raw counts *)
    DIVERT_DELAY : TIME := T#1980ms;    (* eye-to-plate travel, less average polling latency *)
    BELTS_OK_DELAY : TIME := T#1s;      (* run feedback must hold this long to feed boxes *)
    BELTS_OK_TMR : TON;                 (* both belts running, debounced *)
    PE_01_RISE : R_TRIG;                (* tall box arrives at PE_01 *)
    DIVERT_TMR_0 : TON;                 (* eye-to-plate travel timer, divert slot 0 *)
    DIVERT_TMR_1 : TON;                 (* eye-to-plate travel timer, divert slot 1 *)
    DIVERT_TMR_2 : TON;                 (* eye-to-plate travel timer, divert slot 2 *)
    DIVERT_TMR_3 : TON;                 (* eye-to-plate travel timer, divert slot 3 *)
    DIVERT_PEND_0 : BOOL;               (* slot 0 holds a tall box on its way to the pusher *)
    DIVERT_PEND_1 : BOOL;               (* slot 1 holds a tall box on its way to the pusher *)
    DIVERT_PEND_2 : BOOL;               (* slot 2 holds a tall box on its way to the pusher *)
    DIVERT_PEND_3 : BOOL;               (* slot 3 holds a tall box on its way to the pusher *)
    NEXT_SLOT : INT := 0;               (* ring index: the slot the next tall box takes, 0..3 *)
    DIVERT_OVERRUN : BOOL;              (* latched: a tall box found its slot busy and was lost *)
    PUSH_CMD : BOOL;                    (* pusher extend request, held until the extended limit *)
  END_VAR

  (* 1. Belts run at 100 % *)
  CONV_01_RUN_DO := TRUE;
  CONV_02_RUN_DO := TRUE;
  CONV_01_SPD_AO := SPEED_RAW;
  CONV_02_SPD_AO := SPEED_RAW;

  (* 2. Feed boxes only after both belts have reported running for BELTS_OK_DELAY *)
  BELTS_OK_TMR(IN := CONV_01_RUN_DI AND CONV_02_RUN_DI, PT := BELTS_OK_DELAY);
  EMT_01_EN_DO := BELTS_OK_TMR.Q;

  (* 3. Tall box at the eye: give it the next slot and its own travel timer *)
  PE_01_RISE(CLK := PE_01_DI);
  IF PE_01_RISE.Q THEN
    CASE NEXT_SLOT OF
      0: DIVERT_OVERRUN := DIVERT_OVERRUN OR DIVERT_PEND_0; DIVERT_PEND_0 := TRUE;
      1: DIVERT_OVERRUN := DIVERT_OVERRUN OR DIVERT_PEND_1; DIVERT_PEND_1 := TRUE;
      2: DIVERT_OVERRUN := DIVERT_OVERRUN OR DIVERT_PEND_2; DIVERT_PEND_2 := TRUE;
      3: DIVERT_OVERRUN := DIVERT_OVERRUN OR DIVERT_PEND_3; DIVERT_PEND_3 := TRUE;
    END_CASE;
    NEXT_SLOT := (NEXT_SLOT + 1) MOD 4;
  END_IF;

  (* 3a. Each slot's box is due at the plate: extend *)
  DIVERT_TMR_0(IN := DIVERT_PEND_0, PT := DIVERT_DELAY);
  IF DIVERT_TMR_0.Q THEN
    DIVERT_PEND_0 := FALSE;
    PUSH_CMD := TRUE;
  END_IF;
  DIVERT_TMR_1(IN := DIVERT_PEND_1, PT := DIVERT_DELAY);
  IF DIVERT_TMR_1.Q THEN
    DIVERT_PEND_1 := FALSE;
    PUSH_CMD := TRUE;
  END_IF;
  DIVERT_TMR_2(IN := DIVERT_PEND_2, PT := DIVERT_DELAY);
  IF DIVERT_TMR_2.Q THEN
    DIVERT_PEND_2 := FALSE;
    PUSH_CMD := TRUE;
  END_IF;
  DIVERT_TMR_3(IN := DIVERT_PEND_3, PT := DIVERT_DELAY);
  IF DIVERT_TMR_3.Q THEN
    DIVERT_PEND_3 := FALSE;
    PUSH_CMD := TRUE;
  END_IF;

  (* 4. Retract on the extended limit *)
  IF CYL_01_EXT_DI THEN
    PUSH_CMD := FALSE;
  END_IF;
  CYL_01_EXT_DO := PUSH_CMD;
END_PROGRAM

CONFIGURATION Config0
  RESOURCE Res0 ON PLC
    TASK task0(INTERVAL := T#20ms, PRIORITY := 0);
    PROGRAM instance0 WITH task0 : sorter;
  END_RESOURCE
END_CONFIGURATION

(* ---- tank-level-onoff.st ---- *)
(*
  OpenFactory example PLC program: tank-level-onoff (scenes/tank-level-onoff.yaml), the first
  process scene of PLAN 3.3.
  Target: OpenPLC v3 runtime (IEC 61131-3 Structured Text), talking to the OpenFactory simulator
  as a Modbus TCP Slave Device. Setup: docs/guides/openplc-quickstart.md, then
  docs/guides/tank-level-onoff.md for this scene.

  Training and demo use only. Not a safety-rated program and not a safety-rated simulation.

  Sequence of operations
    1. The low level switch (LSL, TK_02_LSL_DI) starts the fill pump P_01.
    2. The pump runs on (seal-in) until the high level switch (LSH, TK_02_LSH_DI) stops it, so the
       level swings between the two switches instead of chattering at one: on/off control with
       the switches as the deadband.
    3. If both switches read on at once (a wiring or switch fault: the tank cannot be both low
       and high), the pump stops.

  I/O map: Modbus addresses come from the scene's int16_scaled lockfile
  (scenes/tank-level-onoff.int16_scaled.modbus.yaml) and the exported I/O list CSV. OpenPLC
  places a Slave Device's points from address 100 onward, so a zero-based Modbus address N maps
  to %IX100.N, %QX100.N, or %IW100+N. TK_02_LT_AI is not used by the sequence; it is there to
  trend or display (raw 0 to 32767 for 0 to 1 m of level).
*)
PROGRAM tank_onoff
  VAR
    (* Discrete inputs from the simulator (Modbus DI:0..3) *)
    P_01_RUN_DI AT %IX100.0 : BOOL;     (* DI:0 Head Tank Fill Pump - running feedback *)
    TK_02_LSH_DI AT %IX100.1 : BOOL;    (* DI:1 Head Tank - high level switch (LSH) *)
    TK_02_LSL_DI AT %IX100.2 : BOOL;    (* DI:2 Head Tank - low level switch (LSL) *)
    SIM_HEARTBEAT_DI AT %IX100.3 : BOOL; (* DI:3 OpenFactory simulator heartbeat, 1 Hz; not used here, watch it for a sim-down watchdog *)
    (* Coils to the simulator (Modbus CO:0) *)
    P_01_RUN_DO AT %QX100.0 : BOOL;     (* CO:0 Head Tank Fill Pump - run command *)
    (* Input registers (Modbus IR:0) *)
    TK_02_LT_AI AT %IW100 : INT;        (* IR:0 Head Tank - level, 0 to 32767 = 0 to 1 m *)
  END_VAR
  VAR
    FILL : BOOL;                        (* the pump is filling (seal-in) *)
  END_VAR

  (* 1-2. Start at low, seal in, stop at high; 3. both switches on is a fault: stop *)
  FILL := (TK_02_LSL_DI OR FILL) AND NOT TK_02_LSH_DI;
  P_01_RUN_DO := FILL;
END_PROGRAM

CONFIGURATION Config0
  RESOURCE Res0 ON PLC
    TASK task0(INTERVAL := T#20ms, PRIORITY := 0);
    PROGRAM instance0 WITH task0 : tank_onoff;
  END_RESOURCE
END_CONFIGURATION

(* ---- tank-level-pid.st ---- *)
(*
  OpenFactory example PLC program: tank-level-pid (scenes/tank-level-pid.yaml), a level loop of
  PLAN 3.3 closed with OpenPLC's PID function block.
  Target: OpenPLC v3 runtime (IEC 61131-3 Structured Text), talking to the OpenFactory simulator
  as a Modbus TCP Slave Device. Setup: docs/guides/openplc-quickstart.md, then
  docs/guides/tank-level-pid.md for this scene.

  Training and demo use only. Not a safety-rated program and not a safety-rated simulation.

  The PID block is the one in OpenPLC's compiler library (matiec lib/pid_st.txt, from the IEC
  61131-3 2nd edition draft): XOUT := KP * (ERROR + ITERM.XOUT / TR + DTERM.XOUT * TD) with
  ERROR := PV - SP. The error is PV minus SP, so a loop that opens the inlet valve on a low level
  needs a negative KP. Its integral (lib/integral_st.txt) is a rectangular sum of ERROR times
  TIME_TO_REAL(CYCLE). It has no output limit and no anti-windup: LIMIT clamps the output here,
  and the interlock holds the block in manual so it cannot wind up while overridden.
  [TBD: verify on the first OpenPLC run] that TIME_TO_REAL(T#20ms) is 0.02 (seconds) in the
  runtime; the gains below assume seconds, as the stand-in script does.

  Sequence of operations
    1. Read the level from the transmitter, raw 0 to 32767 for 0 to 2 m.
    2. PI control: the valve position is KP * (e + sum(e * 0.02 s) / TR) with e = level - 1.0 m.
    3. The output is limited to 0 to 100 % and written to the valve, raw 0 to 32767.
    4. Interlock: while the high level switch (LSH) is on, the valve is closed and the PID is
       held in manual at 0 % (no windup while it is overridden).
    5. For the first second the PID runs in manual at the valve's starting position (66 %),
       tracking the level, then switches to automatic bumplessly: the level input reads 0 until
       its first poll, and starting in automatic on that would slam the valve shut.

  I/O map: Modbus addresses come from the scene's int16_scaled lockfile
  (scenes/tank-level-pid.int16_scaled.modbus.yaml) and the exported I/O list CSV. OpenPLC places
  a Slave Device's points from address 100 onward, so a zero-based Modbus address N maps to
  %IX100.N, %IW100+N, or %QW100+N.
*)
PROGRAM tank_pid
  VAR
    (* Discrete inputs from the simulator (Modbus DI:0..1) *)
    TK_01_LSH_DI AT %IX100.0 : BOOL;    (* DI:0 Level Control Tank - high level switch (LSH), 1.8 m *)
    SIM_HEARTBEAT_DI AT %IX100.1 : BOOL; (* DI:1 OpenFactory simulator heartbeat, 1 Hz; not used here, watch it for a sim-down watchdog *)
    (* Input registers (Modbus IR:0..1) *)
    FV_01_ZT_AI AT %IW100 : INT;        (* IR:0 Tank Inlet Level Control Valve - position feedback, 0 to 32767 = 0 to 100 % *)
    TK_01_LT_AI AT %IW101 : INT;        (* IR:1 Level Control Tank Level Transmitter, 0 to 32767 = 0 to 2 m *)
    (* Holding registers to the simulator (Modbus HR:0) *)
    FV_01_POS_AO AT %QW100 : INT;       (* HR:0 Tank Inlet Level Control Valve - position command, 0 to 32767 = 0 to 100 % *)
  END_VAR
  VAR
    SP : REAL := 1.0;                   (* level setpoint, m *)
    KP : REAL := -400.0;                (* % per m; negative: the PID's error is PV - SP *)
    TR : REAL := 6.0;                   (* reset time, s *)
    START_PCT : REAL := 66.0;           (* valve position at start, % *)
    STARTUP_DELAY : TIME := T#1s;       (* manual until the level reading is live *)
    STARTUP_TMR : TON;
    LIC : PID;                          (* the level controller *)
    LEVEL_M : REAL;
    MANUAL_X0 : REAL;
    OUT_PCT : REAL;
  END_VAR

  (* 1. Level in metres *)
  LEVEL_M := INT_TO_REAL(TK_01_LT_AI) * 2.0 / 32767.0;

  (* 5. Manual at the starting position until the startup delay is done *)
  STARTUP_TMR(IN := TRUE, PT := STARTUP_DELAY);
  IF STARTUP_TMR.Q THEN
    MANUAL_X0 := 0.0;
  ELSE
    MANUAL_X0 := START_PCT / KP;         (* in manual the block outputs KP * X0 *)
  END_IF;

  (* 2. PI on the level; 4. held in manual at 0 % while the high switch overrides it *)
  LIC(AUTO := STARTUP_TMR.Q AND NOT TK_01_LSH_DI, PV := LEVEL_M, SP := SP, X0 := MANUAL_X0,
      KP := KP, TR := TR, TD := 0.0, CYCLE := T#20ms);

  (* 3. Limit to the valve's range; 4. the interlock closes it *)
  IF TK_01_LSH_DI THEN
    OUT_PCT := 0.0;
  ELSE
    OUT_PCT := LIMIT(0.0, LIC.XOUT, 100.0);
  END_IF;
  FV_01_POS_AO := REAL_TO_INT(OUT_PCT * 32767.0 / 100.0);
END_PROGRAM

CONFIGURATION Config0
  RESOURCE Res0 ON PLC
    TASK task0(INTERVAL := T#20ms, PRIORITY := 0);
    PROGRAM instance0 WITH task0 : tank_pid;
  END_RESOURCE
END_CONFIGURATION

(* ---- two-lane-merge.st ---- *)
(*
  OpenFactory example PLC program: two-lane-merge (scenes/two-lane-merge.yaml), PLAN 2.7.
  Target: OpenPLC v3 runtime (IEC 61131-3 Structured Text), talking to the OpenFactory simulator
  as a Modbus TCP Slave Device. Setup: docs/guides/openplc-quickstart.md, then
  docs/guides/two-lane-merge.md for this scene.

  Training and demo use only. Not a safety-rated program and not a safety-rated simulation.

  Sequence of operations
    1. Run both lanes and the outfeed; enable both box sources once all three report running for
       1 s. The lane stoppers are spring-raised (the scene binds raise with invert: true): a
       lane's box waits at its blade until the program energizes STP_x_REL_DO for RELEASE, which
       lets exactly one box through.
    2. STATE 0, idle at 0 degrees with the deck stopped: serve a waiting box (PE_A or PE_B),
       alternating lanes when both wait.
    3. STATE 10, lane A (straight on): release one box and run the deck. The box rides through
       onto the outfeed; the deck is free again when PE_TTA has seen it come and go.
    4. Lane B (from the side): STATE 20 turns the deck to 90; STATE 21, at 90, releases one box
       and runs the deck until PE_TTB sees it centred; STATE 22 stops the deck and turns back;
       STATE 23, at 0, runs the deck until PE_TTA has seen the box come and go.

  Release pulse: the blade takes 0.2 s to drop, and a box at 0.5 m/s is over the blade line for
  0.6 s after that, so a 500 ms pulse ends while the released box is still over the line (it
  passes) and before the next box's front reaches it (it stops). OpenPLC's polling delays both
  edges of the pulse alike, so it does not change the window.

  I/O map: Modbus addresses come from the scene's int16_scaled lockfile
  (scenes/two-lane-merge.int16_scaled.modbus.yaml) and the exported I/O list CSV. OpenPLC places a
  Slave Device's points from address 100 onward, eight bits to a byte: zero-based Modbus address
  N maps to %IX(100 + N / 8).(N MOD 8), so DI:8 is %IX101.0, and likewise for %QX. The scene has
  no analog tags, so both lockfiles give the same addresses.
*)
PROGRAM merge
  VAR
    (* Discrete inputs from the simulator (Modbus DI:0..9) *)
    CONV_A_RUN_DI AT %IX100.0 : BOOL;   (* DI:0 Lane A Infeed Belt Conveyor - running *)
    CONV_B_RUN_DI AT %IX100.1 : BOOL;   (* DI:1 Lane B Infeed Belt Conveyor - running *)
    CONV_OUT_RUN_DI AT %IX100.2 : BOOL; (* DI:2 Merged Outfeed Belt Conveyor - running *)
    PE_A_DI AT %IX100.3 : BOOL;         (* DI:3 Lane A Box Waiting Photo Eye *)
    PE_B_DI AT %IX100.4 : BOOL;         (* DI:4 Lane B Box Waiting Photo Eye *)
    PE_TTA_DI AT %IX100.5 : BOOL;       (* DI:5 Turntable Straight-Through Photo Eye *)
    PE_TTB_DI AT %IX100.6 : BOOL;       (* DI:6 Turntable Side Load Centred Photo Eye *)
    TT_01_AT0_DI AT %IX100.7 : BOOL;    (* DI:7 Lane Merge Turntable - at 0 degrees *)
    TT_01_AT90_DI AT %IX101.0 : BOOL;   (* DI:8 Lane Merge Turntable - at 90 degrees *)
    SIM_HEARTBEAT_DI AT %IX101.1 : BOOL; (* DI:9 OpenFactory simulator heartbeat, 1 Hz; not used here, watch it for a sim-down watchdog *)
    (* Coils to the simulator (Modbus CO:0..8) *)
    CONV_A_RUN_DO AT %QX100.0 : BOOL;   (* CO:0 Lane A Infeed Belt Conveyor - run *)
    CONV_B_RUN_DO AT %QX100.1 : BOOL;   (* CO:1 Lane B Infeed Belt Conveyor - run *)
    CONV_OUT_RUN_DO AT %QX100.2 : BOOL; (* CO:2 Merged Outfeed Belt Conveyor - run *)
    EMT_A_EN_DO AT %QX100.3 : BOOL;     (* CO:3 Lane A Box Source - enable *)
    EMT_B_EN_DO AT %QX100.4 : BOOL;     (* CO:4 Lane B Box Source - enable *)
    STP_A_REL_DO AT %QX100.5 : BOOL;    (* CO:5 Lane A Release Stopper - energize to release *)
    STP_B_REL_DO AT %QX100.6 : BOOL;    (* CO:6 Lane B Release Stopper - energize to release *)
    TT_01_RUN_DO AT %QX100.7 : BOOL;    (* CO:7 Lane Merge Turntable - deck belt run *)
    TT_01_TURN_DO AT %QX101.0 : BOOL;   (* CO:8 Lane Merge Turntable - turn to 90 *)
  END_VAR
  VAR
    BELTS_OK_DELAY : TIME := T#1s;      (* run feedback must hold this long to feed boxes *)
    RELEASE : TIME := T#500ms;          (* stopper release pulse: one box *)
    BELTS_OK_TMR : TON;                 (* lanes and outfeed running, debounced *)
    REL_A_TMR : TON;                    (* lane A stopper energized this long *)
    REL_B_TMR : TON;                    (* lane B stopper energized this long *)
    STATE : INT := 0;                   (* 0 idle, 10 A pass, 20 B turn out, 21 B load, 22 B turn back, 23 B pass *)
    LAST_B : BOOL;                      (* the last box served came from lane B *)
    REL_A : BOOL;                       (* lane A release pulse in progress *)
    REL_B : BOOL;                       (* lane B release pulse in progress *)
    SEEN : BOOL;                        (* PE_TTA has seen the passing box arrive *)
    FEED_OK : BOOL;                     (* belts proven running *)
  END_VAR

  (* 1. Belts run; feed boxes once they have all reported running for BELTS_OK_DELAY *)
  CONV_A_RUN_DO := TRUE;
  CONV_B_RUN_DO := TRUE;
  CONV_OUT_RUN_DO := TRUE;
  BELTS_OK_TMR(IN := CONV_A_RUN_DI AND CONV_B_RUN_DI AND CONV_OUT_RUN_DI, PT := BELTS_OK_DELAY);
  FEED_OK := BELTS_OK_TMR.Q;
  EMT_A_EN_DO := FEED_OK;
  EMT_B_EN_DO := FEED_OK;

  (* 2. Idle at 0: serve a waiting box, alternating when both lanes wait *)
  IF STATE = 0 AND TT_01_AT0_DI THEN
    IF PE_A_DI AND (NOT PE_B_DI OR LAST_B) THEN
      STATE := 10;
      REL_A := TRUE;
      SEEN := FALSE;
      LAST_B := FALSE;
    ELSIF PE_B_DI THEN
      STATE := 20;
      LAST_B := TRUE;
    END_IF;
  END_IF;

  (* 3. Lane A box rides straight through; done when PE_TTA has seen it come and go *)
  IF STATE = 10 THEN
    IF PE_TTA_DI THEN
      SEEN := TRUE;
    ELSIF SEEN THEN
      STATE := 0;
    END_IF;
  END_IF;

  (* 4. Lane B box: turn out, load until centred, turn back, pass through *)
  IF STATE = 20 AND TT_01_AT90_DI THEN
    STATE := 21;
    REL_B := TRUE;
  END_IF;
  IF STATE = 21 AND PE_TTB_DI THEN
    STATE := 22;
  END_IF;
  IF STATE = 22 AND TT_01_AT0_DI THEN
    STATE := 23;
    SEEN := FALSE;
  END_IF;
  IF STATE = 23 THEN
    IF PE_TTA_DI THEN
      SEEN := TRUE;
    ELSIF SEEN THEN
      STATE := 0;
    END_IF;
  END_IF;

  (* Release pulses: one box per pulse *)
  REL_A_TMR(IN := REL_A, PT := RELEASE);
  IF REL_A_TMR.Q THEN
    REL_A := FALSE;
  END_IF;
  REL_B_TMR(IN := REL_B, PT := RELEASE);
  IF REL_B_TMR.Q THEN
    REL_B := FALSE;
  END_IF;
  STP_A_REL_DO := REL_A;
  STP_B_REL_DO := REL_B;
  TT_01_TURN_DO := STATE = 20 OR STATE = 21;
  TT_01_RUN_DO := STATE = 10 OR STATE = 21 OR STATE = 23;
END_PROGRAM

CONFIGURATION Config0
  RESOURCE Res0 ON PLC
    TASK task0(INTERVAL := T#20ms, PRIORITY := 0);
    PROGRAM instance0 WITH task0 : merge;
  END_RESOURCE
END_CONFIGURATION

(* ---- two-tank-cascade.st ---- *)
(*
  OpenFactory example PLC program: two-tank-cascade (scenes/two-tank-cascade.yaml), cascade level
  control of two tanks in series (PLAN 3.3), with two of OpenPLC's PID function blocks.
  Target: OpenPLC v3 runtime (IEC 61131-3 Structured Text), talking to the OpenFactory simulator
  as a Modbus TCP Slave Device. Setup: docs/guides/openplc-quickstart.md, then
  docs/guides/two-tank-cascade.md for this scene.

  Training and demo use only. Not a safety-rated program and not a safety-rated simulation.

  The PID block is the one in OpenPLC's compiler library (matiec lib/pid_st.txt); see
  examples/openplc/tank-level-pid.st for its form. Its error is PV - SP, so both gains are
  negative. It has no output limit or anti-windup: LIMIT clamps both outputs here, and the
  interlock holds both blocks in manual. [TBD: verify on the first OpenPLC run] that
  TIME_TO_REAL(T#20ms) is 0.02 (seconds); the gains assume it, as the stand-in script does.

  Sequence of operations
    1. Read both levels: the upper tank raw 0 to 32767 for 0 to 2 m, the lower for 0 to 1.5 m.
    2. Outer loop (LIC_02): PI on the lower tank's level, setpoint 0.8 m; its output is the upper
       tank's level setpoint, limited to 0.05 to 1.6 m.
    3. Inner loop (LIC_01): PI on the upper tank's level against that setpoint; its output is the
       inlet valve's position, limited to 0 to 100 %.
    4. Interlock: while either tank's high level switch is on, the valve is closed and both
       controllers are held in manual (no windup while they are overridden).
    5. For the first second both controllers run in manual at the plant's starting point (the
       valve at 63 %, the upper level at 0.165 m), then switch to automatic bumplessly. After
       that, the outer block's manual value tracks the upper level, so a return from the
       interlock is bumpless too.

  I/O map: Modbus addresses come from the scene's int16_scaled lockfile
  (scenes/two-tank-cascade.int16_scaled.modbus.yaml) and the exported I/O list CSV. OpenPLC
  places a Slave Device's points from address 100 onward, so a zero-based Modbus address N maps
  to %IX100.N, %IW100+N, or %QW100+N.
*)
PROGRAM tank_cascade
  VAR
    (* Discrete inputs from the simulator (Modbus DI:0..2) *)
    TK_01_LSH_DI AT %IX100.0 : BOOL;    (* DI:0 Upper Tank - high level switch (LSH), 1.8 m *)
    TK_02_LSH_DI AT %IX100.1 : BOOL;    (* DI:1 Lower Tank - high level switch (LSH), 1.35 m *)
    SIM_HEARTBEAT_DI AT %IX100.2 : BOOL; (* DI:2 OpenFactory simulator heartbeat, 1 Hz; not used here, watch it for a sim-down watchdog *)
    (* Input registers (Modbus IR:0..2) *)
    FV_01_ZT_AI AT %IW100 : INT;        (* IR:0 Upper Tank Inlet Control Valve - position feedback, 0 to 100 % *)
    TK_01_LT_AI AT %IW101 : INT;        (* IR:1 Upper Tank Level Transmitter, 0 to 32767 = 0 to 2 m *)
    TK_02_LT_AI AT %IW102 : INT;        (* IR:2 Lower Tank Level Transmitter, 0 to 32767 = 0 to 1.5 m *)
    (* Holding registers to the simulator (Modbus HR:0) *)
    FV_01_POS_AO AT %QW100 : INT;       (* HR:0 Upper Tank Inlet Control Valve - position command, 0 to 100 % *)
  END_VAR
  VAR
    SP2 : REAL := 0.8;                  (* lower tank level setpoint, m *)
    KP_OUTER : REAL := -4.0;            (* m of upper setpoint per m of lower error *)
    TR_OUTER : REAL := 8.0;             (* s *)
    KP_INNER : REAL := -400.0;          (* % per m *)
    TR_INNER : REAL := 3.0;             (* s *)
    UPPER_SP_MIN : REAL := 0.05;        (* m *)
    UPPER_SP_MAX : REAL := 1.6;         (* m *)
    START_PCT : REAL := 63.0;           (* valve position at start, % *)
    START_UPPER : REAL := 0.165;        (* upper level at start, m *)
    STARTUP_DELAY : TIME := T#1s;       (* manual until the level readings are live *)
    STARTUP_TMR : TON;
    LIC_02 : PID;                       (* outer: the lower tank *)
    LIC_01 : PID;                       (* inner: the upper tank *)
    UPPER_M : REAL;
    LOWER_M : REAL;
    HIGH : BOOL;
    AUTO_MODE : BOOL;
    X0_OUTER : REAL;
    X0_INNER : REAL;
    UPPER_SP : REAL;
    OUT_PCT : REAL;
  END_VAR

  (* 1. Levels in metres *)
  UPPER_M := INT_TO_REAL(TK_01_LT_AI) * 2.0 / 32767.0;
  LOWER_M := INT_TO_REAL(TK_02_LT_AI) * 1.5 / 32767.0;
  HIGH := TK_01_LSH_DI OR TK_02_LSH_DI;

  (* 5. Manual at the starting point until the startup delay is done *)
  STARTUP_TMR(IN := TRUE, PT := STARTUP_DELAY);
  AUTO_MODE := STARTUP_TMR.Q AND NOT HIGH;
  IF STARTUP_TMR.Q THEN
    X0_OUTER := UPPER_M / KP_OUTER;      (* in manual the block outputs KP * X0 *)
    X0_INNER := 0.0;
  ELSE
    X0_OUTER := START_UPPER / KP_OUTER;
    X0_INNER := START_PCT / KP_INNER;
  END_IF;

  (* 2. Outer loop: the lower level sets the upper level's setpoint *)
  LIC_02(AUTO := AUTO_MODE, PV := LOWER_M, SP := SP2, X0 := X0_OUTER,
         KP := KP_OUTER, TR := TR_OUTER, TD := 0.0, CYCLE := T#20ms);
  UPPER_SP := LIMIT(UPPER_SP_MIN, LIC_02.XOUT, UPPER_SP_MAX);

  (* 3. Inner loop: the upper level positions the valve *)
  LIC_01(AUTO := AUTO_MODE, PV := UPPER_M, SP := UPPER_SP, X0 := X0_INNER,
         KP := KP_INNER, TR := TR_INNER, TD := 0.0, CYCLE := T#20ms);

  (* 3. Limit to the valve's range; 4. the interlock closes it *)
  IF HIGH THEN
    OUT_PCT := 0.0;
  ELSE
    OUT_PCT := LIMIT(0.0, LIC_01.XOUT, 100.0);
  END_IF;
  FV_01_POS_AO := REAL_TO_INT(OUT_PCT * 32767.0 / 100.0);
END_PROGRAM

CONFIGURATION Config0
  RESOURCE Res0 ON PLC
    TASK task0(INTERVAL := T#20ms, PRIORITY := 0);
    PROGRAM instance0 WITH task0 : tank_cascade;
  END_RESOURCE
END_CONFIGURATION
